(* IEC 61131-3 sources: plc-workbench/experiments/formal_r7/real_model/interlocked_start, 2 files *)

(* ---- candidate_01.st ---- *)
FUNCTION_BLOCK InterlockedStart
VAR_INPUT
  start : BOOL;
  stop : BOOL;
  permit : BOOL;
END_VAR
VAR_OUTPUT
  running : BOOL;
END_VAR
VAR
  prevStart : BOOL;
  startEdge : BOOL;
END_VAR

startEdge := start AND NOT prevStart;
prevStart := start;

IF stop OR NOT permit THEN
  running := FALSE;
ELSIF startEdge THEN
  running := TRUE;
END_IF;
END_FUNCTION_BLOCK

(* ---- candidate_final.st ---- *)
FUNCTION_BLOCK InterlockedStart
VAR_INPUT
  start : BOOL;
  stop : BOOL;
  permit : BOOL;
END_VAR
VAR_OUTPUT
  running : BOOL;
END_VAR
VAR
  prevStart : BOOL;
  startEdge : BOOL;
END_VAR

startEdge := start AND NOT prevStart;
prevStart := start;

IF stop OR NOT permit THEN
  running := FALSE;
ELSIF startEdge THEN
  running := TRUE;
END_IF;
END_FUNCTION_BLOCK
